{attribute 'qualified_only'}
{attribute 'strict'}
TYPE E_PrLine_C_Usage :
(
	eNotInUse := 0,
	eColor_T3,
	eColor_T4
);
END_TYPE

(* stored: Version 1.1.0.1, ProductVersion 3.1.4024.12
   DUT E_PrLine_C_Usage: Id {b16cc458-6e11-4d2b-bb79-bdcfba568582} *)
